// TIA Portal V21 export
// export: Created 2026-10-16T05:44:36.2674366Z, ExportSetting WithDefaults, DisplayName Totally Integrated Automation Portal, DisplayVersion V21 Update 2, DisplayName TIA Portal Test Suite Advanced, DisplayVersion V21, DisplayName SINAMICS Startdrive Advanced, DisplayVersion V21 HF2, DisplayName SINAMICS DCC, DisplayVersion V21, DisplayName SINAMICS Startdrive G110M, G120, G120C, G120D, G120P, G115D, DisplayVersion V21 HF2, DisplayName SINAMICS Startdrive G130, G150, S120, S150, G200, G220, S200, S210, S220, Innomotics MVD, DisplayVersion V21 HF2, DisplayName STEP 7 Professional, DisplayVersion V21 Update 2, DisplayName STEP 7 Safety, DisplayVersion V21, DisplayName Tech WebApplication, DisplayVersion V21, DisplayName WinCC Basic/Comfort/Advanced, DisplayVersion V21 Update 2, DisplayName WinCC Unified, DisplayVersion V21 Update 2
PlcWatchTable "WT05_BoolCreation"
  PlcWatchTableEntry ""TiaMcp_EnableGate_DB".Active"  DisplayFormat=Bool, ModifyTrigger=Permanent, MonitorTrigger=Permanent, Comment="Captured Output state of the selected FB instance: Active"
